{attribute 'pack_mode' := '1'}
TYPE ST_PmsPublish_V1 :
STRUCT
	DeviceIndex			:	UDINT;
	Status				:	UDINT;
	PmsIsAlive			:	UDINT;		// 0: 비정상, 1: 정상
	CpuUsage			:	UDINT;		// %
	CpuTemperature		:	UDINT;		// ℃
	RemainCycle			:	UDINT;		// %
	RemainSaveArea		:	UDINT;		// %
	ProtectModuleCurrent:	REAL;
	ProtectModuleVoltage:	REAL;
	PmsEvent			:	UDINT;
	ModuleStatus1		:	UDINT;
	ModuleStatus2		:	UDINT;
END_STRUCT
END_TYPE

(* stored: Version 1.1.0.1, ProductVersion 3.1.4024.9
   DUT ST_PmsPublish_V1: Id {24fcd318-c2d2-4771-b214-fe565bcf7040} *)
